// TIA Portal V19 export
TYPE "ST_REER_OUTPUT"
   STRUCT
      OUTPUT : Array[0..1] of "ST_Bit";
   END_STRUCT;
END_TYPE
